FUNCTION_BLOCK PID_Level (* Basic Function Block Type *)
  (* Standard: 61499-2 *)
  (* Version 0.0, 5/3/2015, valvya, nxtControl GmbH, Template *)
  PACKAGE Main;
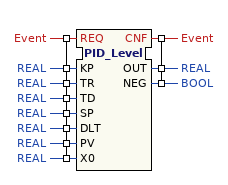
  EVENT_INPUT
    REQ WITH KP, TR, TD, SP, DLT, PV, X0; (* Normal Execution Request *)
  END_EVENT
  EVENT_OUTPUT
    CNF WITH OUT, NEG; (* Execution Confirmation *)
  END_EVENT
  VAR_INPUT
    KP : REAL; (* Input event qualifier *)
    TR : REAL; (* Time in sec *)
    TD : REAL; (* Time in sec *)
    SP : REAL; (* Setpoint *)
    DLT : REAL; (* Time in sec *)
    PV : REAL;
    X0 : REAL;
  END_VAR
  VAR_OUTPUT
    OUT : REAL; (* Output event qualifier *)
    NEG : BOOL;
  END_VAR
  VAR
    ERROR : REAL;
    X1 : REAL;
    X2 : REAL;
    X3 : REAL;
    FIRSTTIME : BOOL := TRUE;
    ITERM : REAL;
    DTERM : REAL;
  END_VAR
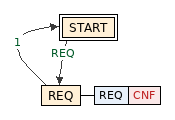
  EC_STATES
    START; (* Initial State *)
    REQ : REQ -> CNF; (* Normal execution *)
  END_STATES
  EC_TRANSITIONS
    START TO REQ := REQ;
    REQ TO START := 1;
  END_TRANSITIONS
  ALGORITHM REQ IN ST: (* PID with Bumpless Transfer and Anti-Reset Windup, REAL PV+XOUT *)
ERROR:=PV-SP;

IF FIRSTTIME THEN
	ITERM:=(ERROR-X0)/KP;
	DTERM:=0;
ELSE
	ITERM:=ITERM+ERROR*DLT/TR;
	DTERM:=(3*(PV-X3)+X1-X2)*TD/DLT/10;
END_IF;
OUT:=-KP*ERROR-ITERM-DTERM;
X3:=X2;X2:=X1;X1:=PV;
ITERM:=ITERM-ERROR*DLT/TR;
NEG:=0;
IF OUT<0 THEN
  NEG := 1;
  // OUT:=0;
ELSIF OUT>450 THEN
  OUT:=100;
END_IF;
FIRSTTIME:=FALSE;
  END_ALGORITHM
END_FUNCTION_BLOCK
